(* IEC 61131-3 sources: bcs-engineering-dsl/language/test/generating/switch_test/expected, 4 files *)

(* ---- OperationMode.st ---- *)
{attribute 'qualified_only'}
{attribute 'strict'}
TYPE OperationMode :
(
    IDLE := 0,
    HEATING := 1,
    COOLING := 2,
    ERROR := 3
);
END_TYPE

(* ---- SwitchFB_decl.st ---- *)
FUNCTION_BLOCK SwitchFB
VAR_INPUT
    iMode: OperationMode;
    iTemperature: REAL;
END_VAR
VAR_OUTPUT
    oHeatingValue: REAL;
    oCoolingValue: REAL;
    oStatusMessage: STRING;
END_VAR
VAR
    adjustedTemp: REAL;
END_VAR

(* ---- MAIN_decl.st ---- *)
PROGRAM MAIN
VAR
    TestSwitch_mode: OperationMode := OperationMode.HEATING;
    TestSwitch_temperature: REAL := 22.5;
    TestSwitch_heatingValue: REAL;
    TestSwitch_coolingValue: REAL;
    TestSwitch_statusMsg: STRING;
    SwitchFBInstance1: SwitchFB;
END_VAR

(* ---- SwitchFB_impl.st ---- *)
adjustedTemp := iTemperature * 1.05;
CASE iMode OF
    OperationMode.IDLE:
        oHeatingValue := 0;
        oCoolingValue := 0;
        oStatusMessage := 'System idle';
    OperationMode.HEATING:
        oHeatingValue := adjustedTemp;
        oCoolingValue := 0;
        oStatusMessage := 'Heating active';
    OperationMode.COOLING:
        oHeatingValue := 0;
        oCoolingValue := adjustedTemp;
        oStatusMessage := 'Cooling active';
    ELSE
        oHeatingValue := 0;
        oCoolingValue := 0;
        oStatusMessage := 'Error state';
END_CASE;
